SUBAPPLICATION AS_GT_0 (* Prüft ob SINT-Adapter Wert > 0 ist (AX-Adapter Ausgang) *)
  (* Standard: 61499-2 *)
  (* Version 1.0, 2026-10-15, franz, Meisterschulen am Ostbahnhof *)
  PACKAGE MyLib::sys;
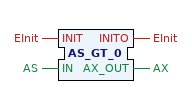
  EVENT_INPUT
    INIT : EInit; (* Initialization Request *)
  END_EVENT
  EVENT_OUTPUT
    INITO : EInit; (* Initialization Confirm *)
  END_EVENT
  SOCKETS
    IN : adapter::types::unidirectional::AS;
  END_SOCKETS
  PLUGS
    AX_OUT : adapter::types::unidirectional::AX;
  END_PLUGS
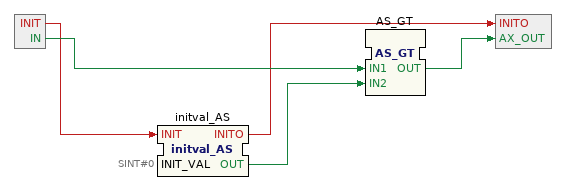
  FBS
    AS_GT : adapter::iec61131::comparison::AS_GT;
    initval_AS : adapter::types::unidirectional::AS::initval::initval_AS(INIT_VAL := SINT#0);
  END_FBS
  EVENT_CONNECTIONS
    INIT TO initval_AS.INIT;
    initval_AS.INITO TO INITO;
  END_CONNECTIONS
  ADAPTER_CONNECTIONS
    IN TO AS_GT.IN1;
    AS_GT.OUT TO AX_OUT;
    initval_AS.OUT TO AS_GT.IN2;
  END_CONNECTIONS
END_SUBAPPLICATION
